// TIA Portal V20 export
Screen "SEW_FIFO"  1276x673
  ScreenItem "Title_ScreenOverview_X390_Y2" at 390,7 size 510x57  Type=HmiTextBox
  ScreenItem "符号 IO 域_7" at 479,72 size 290x38  Type=HmiSymbolicIOField
  ScreenItem "permanentareaborderrectangle" at 0,0 size 0x0  Type=HmiRectangle
  ScreenItem "Line_Header_X0_Y64" at 0,65 size 1276x0  Type=HmiLine
  ScreenItem "Button_Back" at 2,2 size 90x60  Type=HmiButton
  ScreenItem "Faceplate container_1" at 0,110 size 1276x547  Type=HmiFaceplateContainer
